Fanuc KAREL source: kt00298.KL

-- PROVISIONAL review KL for V1013-1; original PC SHA256 384d87ffee2e710ebf029584dcb4e8aa55432529aa8657ab385a99b3211f18c6
-- Incomplete behavior may be omitted. Consult companion uncertainty JSON. Do not deploy.
PROGRAM KT00298
%NOLOCKGROUP
VAR
  R1 : REAL
  R2 : REAL
  OUT : BOOLEAN
BEGIN
  -- UNRESOLVED_PC offsets 5-16; opcodes 2E,23
  -- UNRESOLVED_PC offsets 21-32; opcodes 2E,23
  -- UNRESOLVED_PC offsets 37-48; opcodes 2E,23
  -- UNRESOLVED_PC offsets 53-64; opcodes 2E,23
  -- UNRESOLVED_PC offsets 69-88; opcodes 21,21,6E,23
  -- UNRESOLVED_PC offsets 93-97; opcodes 7F
END KT00298
